Fanuc KAREL source: KD00072.KL

PROGRAM KD00072
%NOLOCKGROUP
VAR
  I: INTEGER
  J: INTEGER
  B: BOOLEAN
  R: REAL
  S: STRING[80]
BEGIN
  PULSE DOUT[1] FOR 100 NOWAIT
END KD00072
